# EPICS autosave request: iocs/quadem/db/quadEM_TimeSeries_settings.req
# FILE... quadEM_TimeSeries_settings.req
$(P)$(R)ReadAll.SCAN
$(P)$(R)NuseAll
$(P)$(R)Dwell
$(P)$(R)PresetReal
$(P)$(R)AutoRestartTS
$(P)$(R)ComputeFFT
$(P)$(R)EnableClientWait
